Fanuc KAREL source: kb00046.KL

-- PROVISIONAL review KL for V770-1; original PC SHA256 c193e5887b2e2089dec023ace6c93da0bcd75d5140e6d9a89e1530287e639a6e
-- Incomplete behavior may be omitted. Consult companion uncertainty JSON. Do not deploy.
PROGRAM KB00046
%NOLOCKGROUP
BEGIN
  -- UNRESOLVED_PC offsets 5-14; opcodes 3F,75
  -- UNRESOLVED_PC offsets 19-28; opcodes 3F,75
  -- UNRESOLVED_PC offsets 33-40; opcodes 9D,23
  -- UNRESOLVED_PC offsets 45-52; opcodes 9D,23
  -- UNRESOLVED_PC offsets 57-64; opcodes 9D,23
  -- UNRESOLVED_PC offsets 69-107; opcodes 27,22,2A,22,2A,22,22,22,31
  -- UNRESOLVED_PC offsets 112-116; opcodes 7F
END KB00046
